(* IEC 61131-3 sources: SemaPLC/sema-plc-benchmark/spec2control-benchmark/data/st-baseline/paper-machine/pous/programs, 10 files *)

(* ---- main.st ---- *)
PROGRAM main
VAR
	Heartbeat : bool;
END_VAR

(* Entry point required by OpenPLC Editor v4. The process sections run as parallel program instances under task0; main only provides a scan heartbeat. *)
Heartbeat := NOT Heartbeat;

END_PROGRAM

(* ---- Section10.st ---- *)
PROGRAM Section10
VAR
	FT901_NipLoad_kN : real;
	FT902_FlowRate_Lmin : real;
	FIC904_Flow_SP_FromRatio : real;
	FT_901 : ANALOG_IN;
	FT_902 : ANALOG_IN;
	CW_901 : ANALOG_IN;
	FFIC_903 : RATIO_CONTROL;
	FIC_904 : PID_BASIC;
	FV_104 : VALVE_ELECTRIC;
	XV_105 : VALVE_ON_OFF;
	NipLoadOK_NOT : bool;
	SP_LowCut_SEL : real;
	XV105Closed_NOT : bool;
	CW901DevTrip_OR : bool;
	FT901_LowOrFault_OR : bool;
	CW901_DevOrFault_OR : bool;
	Interlock_PermissivesFail1_OR : bool;
	Interlock_PermissivesFail2_OR : bool;
	FFIC903_Inhibit_OR : bool;
END_VAR

FT_901(
    PV_Low := 5.0,
    Scaling_Slope := 6.25,
    Scaling_Offset := -25.0,
    Alarm_Enable := TRUE);
FT_902(
    Scaling_Slope := 31.25,
    Scaling_Offset := -125.0,
    Alarm_Enable := TRUE);
CW_901(
    Alarm_Enable := TRUE);
FT901_LowOrFault_OR := FT_901.Low_Alarm OR FT_901.General_Fault;
XV_105();
XV105Closed_NOT := NOT XV_105.FB_Opened;
Interlock_PermissivesFail1_OR := XV105Closed_NOT OR FT901_LowOrFault_OR;
CW901DevTrip_OR := CW_901.High_Alarm OR CW_901.Low_Alarm;
CW901_DevOrFault_OR := CW901DevTrip_OR OR CW_901.General_Fault;
Interlock_PermissivesFail2_OR := FT_902.General_Fault OR CW901_DevOrFault_OR;
FFIC903_Inhibit_OR := Interlock_PermissivesFail1_OR OR Interlock_PermissivesFail2_OR;
FFIC_903(
    Auto := TRUE,
    PrimaryPV := FT_901.PV,
    SecondaryPV := FT_902.PV,
    RatioSP := 2.0,
    Bias := 0.0,
    MV_MIN := 0.0,
    MV_MAX := 500.0,
    Inhibit := FFIC903_Inhibit_OR);
NipLoadOK_NOT := NOT FT_901.Low_Alarm;
SP_LowCut_SEL := SEL(G := NipLoadOK_NOT, IN0 := 0.0, IN1 := FFIC_903.SlaveSP);
FIC_904(
    AUTO := TRUE,
    PV := FT_902.PV,
    SP := SP_LowCut_SEL,
    MV_MIN := 0.0,
    MV_MAX := 100.0,
    X0 := 0.0,
    Deviation_Limit := 5.0);
FV_104(
    Control_Signal := FIC_904.XOUT,
    Manual_Mode := FALSE,
    Open_Limit := 100.0,
    Close_Limit := 0.0,
    Inhibit := FFIC903_Inhibit_OR);

(* Outputs published to other sections / HMI. *)
FT901_NipLoad_kN := FT_901.PV;
FT902_FlowRate_Lmin := FT_902.PV;
FIC904_Flow_SP_FromRatio := FFIC_903.SlaveSP;

END_PROGRAM

(* ---- Section2.st ---- *)
PROGRAM Section2
VAR
	LT_101_Flow_PV : real;
	FC_101_MV_to_FV106 : real;
	M_102_VSD_Speed_Out : real;
	Flow_Deviation_Alarm_30s : bool;
	Flow_High_Alarm : bool;
	Flow_Low_Alarm : bool;
	M_102_Start_Request : bool;
	M_102_Stop_Request : bool;
	LT_101 : ANALOG_IN;
	FC_101 : PID_BASIC;
	M_102 : MOTOR_VSD;
	FV_106 : VALVE_ELECTRIC;
	LV_103 : VALVE_ELECTRIC;
	XV_102 : VALVE_ON_OFF;
	XV_104 : VALVE_ON_OFF;
	XV_105 : VALVE_ON_OFF;
	FlowDeviationAlarm_TON : TON;
	M102_RestartDelay_TON : TON;
	FC101_ValvesOpen_AND : bool;
	FC101_ValvesNotOpen_NOT : bool;
	FC101_Inhibit_OR : bool;
	M102_XV105NotClosed_NOT : bool;
	M102_Inhibit_OR : bool;
	M102_InhibitNot_NOT : bool;
	M102_StartPermissive_AND : bool;
	M102_StopCmd_OR : bool;
	HopperLevelAbove20_GT : bool;
END_VAR

LT_101(
    PV_High := 380.0,
    PV_Low := 20.0,
    Scaling_Slope := 25.0,
    Scaling_Offset := -100.0,
    Alarm_Enable := TRUE);
XV_105(
    Timeout := T#5s);
M102_XV105NotClosed_NOT := NOT XV_105.FB_Closed;
M102_Inhibit_OR := M102_XV105NotClosed_NOT OR LT_101.General_Fault;
LV_103(
    Open_Limit := 100.0,
    Close_Limit := 0.0);
HopperLevelAbove20_GT := (LV_103.Feedback_Pos > 20.0);
M102_InhibitNot_NOT := NOT M102_Inhibit_OR;
M102_RestartDelay_TON(
    IN := M102_InhibitNot_NOT,
    PT := T#60s);
M102_StartPermissive_AND := HopperLevelAbove20_GT AND XV_105.FB_Closed AND M102_RestartDelay_TON.Q AND M_102_Start_Request;
M102_StopCmd_OR := M_102_Stop_Request OR M102_Inhibit_OR;
M_102(
    Start_Cmd := M102_StartPermissive_AND,
    Stop_Cmd := M102_StopCmd_OR,
    Accel_Ramp := T#2s,
    Decel_Ramp := T#2s,
    Inhibit := M102_Inhibit_OR);
XV_102(
    Timeout := T#5s,
    Inhibit := M_102.FB_Fault);
XV_104(
    Timeout := T#5s,
    Inhibit := M_102.FB_Fault);
FC101_ValvesOpen_AND := XV_102.FB_Opened AND XV_104.FB_Opened;
FC101_ValvesNotOpen_NOT := NOT FC101_ValvesOpen_AND;
FC101_Inhibit_OR := FC101_ValvesNotOpen_NOT OR LT_101.General_Fault OR M_102.FB_Fault;
FC_101(
    AUTO := TRUE,
    PV := LT_101.PV,
    SP := 250.0,
    MV_MIN := 0.0,
    MV_MAX := 100.0,
    KP := 3.0,
    TR := 1.2,
    TD := 0.3,
    Deviation_Limit := 5.0,
    Inhibit := FC101_Inhibit_OR);
FV_106(
    Control_Signal := FC_101.XOUT,
    Manual_Mode := FALSE,
    Manual_Position := 0.0,
    Open_Limit := 100.0,
    Close_Limit := 0.0,
    Timeout := T#5s,
    Inhibit := LT_101.General_Fault);
FlowDeviationAlarm_TON(
    IN := FC_101.Deviation_Alarm,
    PT := T#30s);

(* Outputs published to other sections / HMI. *)
FC_101_MV_to_FV106 := FC_101.XOUT;
LT_101_Flow_PV := LT_101.PV;
Flow_High_Alarm := LT_101.High_Alarm;
Flow_Low_Alarm := LT_101.Low_Alarm;
Flow_Deviation_Alarm_30s := FlowDeviationAlarm_TON.Q;
M_102_VSD_Speed_Out := M_102.Speed_Out;

END_PROGRAM

(* ---- Section3.st ---- *)
PROGRAM Section3
VAR
	TT_103_Temperature_PV : real;
	PT_101_Pressure_PV : real;
	TIC_104_RSP_to_FC_203 : real;
	PIC_101_RSP_to_FC_202 : real;
	FC_203_MV_to_SV_203 : real;
	FC_202_MV_to_FV_202 : real;
	TT_103 : ANALOG_IN;
	PT_101 : ANALOG_IN;
	TIC_104 : PID_BASIC;
	PIC_101 : PID_BASIC;
	FC_203 : PID_BASIC;
	FC_202 : PID_BASIC;
	SV_203 : VALVE_ELECTRIC;
	FV_202 : VALVE_ELECTRIC;
	SV203Trip_OR : bool;
	CascadeInhibit_OR : bool;
END_VAR

TT_103(
    PV_High := 180.0,
    PV_Low := 160.0,
    Scaling_Slope := 11.25,
    Scaling_Offset := -25.0,
    Alarm_Enable := TRUE);
PT_101(
    Alarm_Enable := TRUE);
PIC_101(
    AUTO := TRUE,
    PV := PT_101.PV,
    SP := 800.0,
    MV_MIN := 0.0,
    MV_MAX := 100.0,
    PV_High := 850.0,
    PV_Low := 750.0,
    Inhibit := CascadeInhibit_OR);
FC_202(
    AUTO := TRUE,
    SP := PIC_101.XOUT,
    MV_MIN := 0.0,
    MV_MAX := 100.0,
    Inhibit := PIC_101.PV_Low_Alarm);
FV_202(
    Control_Signal := FC_202.XOUT);
FC_203(
    AUTO := TRUE,
    SP := TIC_104.XOUT,
    MV_MIN := 0.0,
    MV_MAX := 100.0,
    KP := 3.5,
    TR := 0.3,
    Inhibit := TT_103.General_Fault);
SV203Trip_OR := PIC_101.PV_High_Alarm OR TIC_104.PV_High_Alarm;
SV_203(
    Control_Signal := FC_203.XOUT,
    Inhibit := SV203Trip_OR);
CascadeInhibit_OR := TT_103.General_Fault OR PT_101.General_Fault OR SV_203.Alarm OR FV_202.Alarm;
TIC_104(
    AUTO := TRUE,
    PV := TT_103.PV,
    SP := 170.0,
    MV_MIN := 0.0,
    MV_MAX := 100.0,
    KP := 1.2,
    TR := 2.0,
    Inhibit := CascadeInhibit_OR);

(* Outputs published to other sections / HMI. *)
TT_103_Temperature_PV := TT_103.PV;
PT_101_Pressure_PV := PT_101.PV;
TIC_104_RSP_to_FC_203 := TIC_104.XOUT;
PIC_101_RSP_to_FC_202 := PIC_101.XOUT;
FC_203_MV_to_SV_203 := FC_203.XOUT;
FC_202_MV_to_FV_202 := FC_202.XOUT;

END_PROGRAM

(* ---- Section4.st ---- *)
PROGRAM Section4
VAR
	PIT103_Pressure_kPa : real;
	PT101_UpstreamPressure_kPa : real;
	DT301_PulpDensity_Pct : real;
	PIC104_ControlOutput_to_FV106_Pct : real;
	FV106_ValvePositionFeedback_Pct : real;
	DT_301 : ANALOG_IN;
	PIT_103 : ANALOG_IN;
	PT_101 : ANALOG_IN;
	PIC_104 : PID_BASIC;
	FV_106 : VALVE_ELECTRIC;
	XV_102 : VALVE_ON_OFF;
	XV_107 : VALVE_ON_OFF;
	XV_102_OPEN_FB : DIGITAL_IN;
	XV_107_OPEN_FB : DIGITAL_IN;
	PERM_XV102_OPEN : BOOL_INPUT;
	PERM_XV107_OPEN : BOOL_INPUT;
	PIC104Inhibit_OR : bool;
	FV106Inhibit_OR : bool;
	SystemFault_OR : bool;
	XV102NotOpen_NOT : bool;
	XV107NotOpen_NOT : bool;
	SystemEnable_NOT : bool;
	PIC104Auto_NOT : bool;
END_VAR

DT_301();
PIT_103(
    Scaling_Slope := 31.25,
    Scaling_Offset := -125.0);
PT_101();
PIC104Inhibit_OR := PT_101.Low_Alarm OR PT_101.High_Alarm OR DT_301.High_Alarm OR PIT_103.General_Fault;
PIC104Auto_NOT := NOT PIC104Inhibit_OR;
PIC_104(
    AUTO := PIC104Auto_NOT,
    PV := PIT_103.PV,
    SP := 250.0,
    MV_MIN := 0.0,
    MV_MAX := 100.0,
    X0 := 0.0,
    KP := -3.0,
    TR := 1.2,
    TD := 0.1,
    PV_High := 275.0,
    PV_Low := 200.0,
    Deviation_Limit := 12.5,
    Inhibit := PIC104Inhibit_OR);
XV_102_OPEN_FB();
PERM_XV102_OPEN(
    Bool_In := XV_102_OPEN_FB.DI_Out);
XV102NotOpen_NOT := NOT PERM_XV102_OPEN.Bool_Out;
XV_107_OPEN_FB();
PERM_XV107_OPEN(
    Bool_In := XV_107_OPEN_FB.DI_Out);
XV107NotOpen_NOT := NOT PERM_XV107_OPEN.Bool_Out;
FV106Inhibit_OR := XV102NotOpen_NOT OR XV107NotOpen_NOT OR PT_101.High_Alarm OR PIT_103.General_Fault;
FV_106(
    Control_Signal := PIC_104.XOUT,
    Manual_Mode := FALSE,
    Manual_Position := 0.0,
    Open_Limit := 100.0,
    Close_Limit := 0.0,
    Timeout := T#2S,
    Inhibit := FV106Inhibit_OR);
SystemFault_OR := PT_101.General_Fault OR DT_301.General_Fault;
SystemEnable_NOT := NOT SystemFault_OR;
XV_102(
    Open_Cmd := SystemEnable_NOT,
    Close_Cmd := SystemFault_OR,
    Inhibit := SystemFault_OR);
XV_107(
    Open_Cmd := SystemEnable_NOT,
    Close_Cmd := SystemFault_OR,
    Inhibit := SystemFault_OR);

(* Outputs published to other sections / HMI. *)
PIT103_Pressure_kPa := PIT_103.PV;
PT101_UpstreamPressure_kPa := PT_101.PV;
DT301_PulpDensity_Pct := DT_301.PV;
PIC104_ControlOutput_to_FV106_Pct := PIC_104.XOUT;
FV106_ValvePositionFeedback_Pct := FV_106.Feedback_Pos;

END_PROGRAM

(* ---- Section5.st ---- *)
PROGRAM Section5
VAR
	AT102_pH_PV : real;
	AT107_pH_PV : real;
	TIT106_Temperature_PV : real;
	LIC102_MV_to_FV101 : real;
	TIC106_MV_to_FV103 : real;
	LIC104_MV_to_XV104 : real;
	AT_102 : ANALOG_IN;
	AT_107 : ANALOG_IN;
	TIT_106 : ANALOG_IN;
	LIC_102 : PID_BASIC;
	TIC_106 : PID_BASIC;
	LIC_104 : PID_BASIC;
	FV_101 : VALVE_ELECTRIC;
	FV_103 : VALVE_ELECTRIC;
	XV_104 : VALVE_ELECTRIC;
	PHExtremeTrip_OR : bool;
END_VAR

AT_102(
    Scaling_Slope := 0.875,
    Scaling_Offset := -3.5,
    Alarm_Enable := TRUE);
AT_107(
    Alarm_Enable := TRUE);
TIT_106(
    Scaling_Slope := 6.25,
    Scaling_Offset := -25.0,
    Alarm_Enable := TRUE);
FV_101(
    Control_Signal := LIC_102.XOUT,
    Open_Limit := 100.0,
    Close_Limit := 0.0,
    Timeout := T#10s,
    Inhibit := AT_107.General_Fault);
PHExtremeTrip_OR := LIC_102.PV_High_Alarm OR LIC_102.PV_Low_Alarm;
LIC_102(
    AUTO := TRUE,
    PV := AT_102.PV,
    SP := 9.25,
    MV_MIN := 10.0,
    MV_MAX := 90.0,
    X0 := FV_101.Feedback_Pos,
    KP := 1.8,
    TR := 0.5,
    TD := 0.1,
    PV_High := 10.5,
    PV_Low := 8.5,
    Deviation_Limit := 1.0,
    Inhibit := PHExtremeTrip_OR);
FV_103(
    Control_Signal := TIC_106.XOUT,
    Open_Limit := 100.0,
    Close_Limit := 0.0,
    Timeout := T#10s);
TIC_106(
    AUTO := TRUE,
    PV := TIT_106.PV,
    SP := 65.0,
    MV_MIN := 0.0,
    MV_MAX := 100.0,
    X0 := FV_103.Feedback_Pos,
    KP := 2.0,
    TR := 0.4,
    TD := 0.05,
    PV_High := 75.0,
    PV_Low := 55.0,
    Inhibit := TIC_106.PV_High_Alarm);
XV_104(
    Control_Signal := LIC_104.XOUT,
    Open_Limit := 100.0,
    Close_Limit := 0.0,
    Timeout := T#10s);
LIC_104(
    AUTO := TRUE,
    SP := 120.0,
    MV_MIN := 0.0,
    MV_MAX := 100.0,
    X0 := XV_104.Feedback_Pos,
    KP := 1.5,
    TR := 1.0,
    TD := 0.2,
    Deviation_Limit := 10.0);

(* Outputs published to other sections / HMI. *)
AT102_pH_PV := AT_102.PV;
AT107_pH_PV := AT_107.PV;
TIT106_Temperature_PV := TIT_106.PV;
LIC102_MV_to_FV101 := LIC_102.XOUT;
TIC106_MV_to_FV103 := TIC_106.XOUT;
LIC104_MV_to_XV104 := LIC_104.XOUT;

END_PROGRAM

(* ---- Section6.st ---- *)
PROGRAM Section6
VAR
	CT501_Consistency_PV_Pct : real;
	FC502_MV_to_FV502_Pct : real;
	SELT501_SEL_PV_WsPerMm2 : real;
	SELC501_MV_to_PGA501_Pct : real;
	LT501_Level_PV_Pct : real;
	PT502_Pressure_PV_kPa : real;
	PGT501_PlateGap_PV_mm : real;
	CT_501 : ANALOG_IN;
	FC_502 : PID_BASIC;
	FV_502 : VALVE_ELECTRIC;
	LT_501 : ANALOG_IN;
	M_501 : MOTOR_ON_OFF;
	PT_502 : ANALOG_IN;
	SELC_501 : PID_BASIC;
	PGT_501 : ANALOG_IN;
	PGA_501 : VALVE_ELECTRIC;
	SELT_501 : ANALOG_IN;
	INTLK_M501_RUNNING : BOOL_INPUT;
	INTLK_PLATE_GAP_IN_RANGE : BOOL_INPUT;
	INTLK_LEVEL_ABOVE_20 : BOOL_INPUT;
	PERM_PT502_IN_RANGE : BOOL_INPUT;
	PGT501_OutOfRange_OR : bool;
	PlateGapInRange_NOT : bool;
	SEL_Enable_AND : bool;
	SEL_Inhibit_NOT : bool;
	LT501_LevelNotOK_OR : bool;
	LevelAbove20_NOT : bool;
	PT502_NotInRange_OR : bool;
	PT502_InRange_NOT : bool;
	FC502_Inhibit_OR : bool;
END_VAR

CT_501(
    Scaling_Slope := 0.1875,
    Scaling_Offset := 1.25,
    Alarm_Enable := TRUE);
LT_501(
    Alarm_Enable := TRUE);
LT501_LevelNotOK_OR := LT_501.Low_Alarm OR LT_501.General_Fault;
PT_502(
    Alarm_Enable := TRUE);
PT502_NotInRange_OR := PT_502.High_Alarm OR PT_502.Low_Alarm OR PT_502.General_Fault;
FC502_Inhibit_OR := LT501_LevelNotOK_OR OR PT502_NotInRange_OR OR CT_501.General_Fault;
FC_502(
    AUTO := TRUE,
    PV := CT_501.PV,
    SP := 3.0,
    MV_MIN := 0.0,
    MV_MAX := 100.0,
    X0 := 0.0,
    KP := 2.2,
    TR := 0.7,
    TD := 0.0,
    PV_High := 4.0,
    PV_Low := 2.0,
    Inhibit := FC502_Inhibit_OR);
FV_502(
    Control_Signal := FC_502.XOUT,
    Manual_Mode := FALSE,
    Open_Limit := 100.0,
    Close_Limit := 0.0,
    Inhibit := FC502_Inhibit_OR);
PGT_501(
    Alarm_Enable := TRUE);
PGT501_OutOfRange_OR := PGT_501.High_Alarm OR PGT_501.Low_Alarm OR PGT_501.General_Fault;
M_501(
    Inhibit := PGT501_OutOfRange_OR);
SELT_501(
    Scaling_Slope := 0.0625,
    Scaling_Offset := -0.05,
    Alarm_Enable := TRUE);
INTLK_M501_RUNNING(
    Bool_In := M_501.FB_Running);
PlateGapInRange_NOT := NOT PGT501_OutOfRange_OR;
INTLK_PLATE_GAP_IN_RANGE(
    Bool_In := PlateGapInRange_NOT);
SEL_Enable_AND := INTLK_M501_RUNNING.Bool_Out AND INTLK_PLATE_GAP_IN_RANGE.Bool_Out;
SEL_Inhibit_NOT := NOT SEL_Enable_AND;
SELC_501(
    AUTO := TRUE,
    PV := SELT_501.PV,
    MV_MIN := 0.0,
    MV_MAX := 100.0,
    X0 := 0.0,
    KP := 1.8,
    TR := 0.5,
    TD := 0.1,
    PV_High := 1.1,
    PV_Low := 0.3,
    Inhibit := SEL_Inhibit_NOT);
PGA_501(
    Control_Signal := SELC_501.XOUT,
    Manual_Mode := FALSE,
    Open_Limit := 100.0,
    Close_Limit := 0.0);
LevelAbove20_NOT := NOT LT501_LevelNotOK_OR;
INTLK_LEVEL_ABOVE_20(
    Bool_In := LevelAbove20_NOT);
PT502_InRange_NOT := NOT PT502_NotInRange_OR;
PERM_PT502_IN_RANGE(
    Bool_In := PT502_InRange_NOT);

(* Outputs published to other sections / HMI. *)
CT501_Consistency_PV_Pct := CT_501.PV;
FC502_MV_to_FV502_Pct := FC_502.XOUT;
SELT501_SEL_PV_WsPerMm2 := SELT_501.PV;
SELC501_MV_to_PGA501_Pct := SELC_501.XOUT;
LT501_Level_PV_Pct := LT_501.PV;
PT502_Pressure_PV_kPa := PT_502.PV;
PGT501_PlateGap_PV_mm := PGT_501.PV;

END_PROGRAM

(* ---- Section7.st ---- *)
PROGRAM Section7
VAR
	CT_601_PV : real;
	FT_601_PV : real;
	FT_601_SP : real;
	PIT_601_PV : real;
	VT_601_PV : real;
	FS_601_MinFlow_OK : bool;
	P_601_Run_OK : bool;
	FFIC601_Bias : real;
	ALM_601 : bool;
	ALM_601_High : bool;
	ALM_601_Low : bool;
	ALM_602 : bool;
	ALM_603 : bool;
	ALM_604 : bool;
	Process_Permissives_OK : bool;
	MasterInhibit : bool;
	CT601_RateHigh : bool;
	CT_601 : ANALOG_IN;
	FT_601 : ANALOG_IN;
	PIT_601 : ANALOG_IN;
	VT_601 : ANALOG_IN;
	FS_601 : BOOL_INPUT;
	P_601_RUN : BOOL_INPUT;
	FV_601 : VALVE_ELECTRIC;
	FIC_601 : PID_BASIC;
	FFIC_601 : RATIO_CONTROL;
	ProcessUpset_Timer : TON;
	PumpRun_Fault : bool;
	MinFlow_Fault : bool;
	CT_Failure : bool;
	FT_Failure : bool;
	Inhibit_Any : bool;
	Auto_Enable : bool;
	SlaveSP_TooHigh : bool;
	SlaveSP_TooLow : bool;
	SlaveSP_LimitAlarm : bool;
END_VAR

CT_601(
    Alarm_Enable := TRUE);
FT_601(
    PV_High := 500.0,
    PV_Low := 10.0,
    Alarm_Enable := TRUE);
PIT_601(
    PV_Low := 300.0,
    Alarm_Enable := TRUE);
VT_601(
    Alarm_Enable := TRUE);
FS_601(
    Alarm_OnFalse := TRUE);
P_601_RUN(
    Alarm_OnFalse := TRUE);
CT_Failure := CT_601.High_Alarm OR CT_601.Low_Alarm OR CT_601.General_Fault;
FT_Failure := FT_601.High_Alarm OR FT_601.Low_Alarm OR FT_601.General_Fault;
MinFlow_Fault := NOT FS_601.Bool_Out;
PumpRun_Fault := NOT P_601_RUN.Bool_Out;
Inhibit_Any := PumpRun_Fault OR MinFlow_Fault OR PIT_601.Low_Alarm OR VT_601.Low_Alarm OR CT_Failure OR FT_Failure;
Auto_Enable := NOT Inhibit_Any;
FFIC_601(
    Auto := Auto_Enable,
    PrimaryPV := CT_601.PV,
    SecondaryPV := FT_601.PV,
    RatioSP := 2.5,
    Bias := FFIC601_Bias,
    TrimKp := 0.1,
    TrimTi := T#2s,
    MV_MIN := 10.0,
    MV_MAX := 500.0,
    Inhibit := Inhibit_Any);
FIC_601(
    AUTO := Auto_Enable,
    PV := FT_601.PV,
    SP := FFIC_601.SlaveSP,
    MV_MIN := 0.0,
    MV_MAX := 100.0,
    X0 := 20.0,
    Inhibit := Inhibit_Any);
FV_601(
    Control_Signal := FIC_601.XOUT,
    Manual_Mode := Inhibit_Any,
    Manual_Position := 20.0,
    Open_Limit := 100.0,
    Close_Limit := 0.0,
    Inhibit := Inhibit_Any);
ProcessUpset_Timer(
    IN := CT601_RateHigh,
    PT := T#10s);
SlaveSP_TooHigh := (FFIC_601.SlaveSP > 500.0);
SlaveSP_TooLow := (FFIC_601.SlaveSP < 10.0);
SlaveSP_LimitAlarm := SlaveSP_TooHigh OR SlaveSP_TooLow;

(* Outputs published to other sections / HMI. *)
ALM_601 := SlaveSP_LimitAlarm;
ALM_602 := CT_Failure;
ALM_603 := FT_Failure;
ALM_604 := ProcessUpset_Timer.Q;
CT_601_PV := CT_601.PV;
FT_601_PV := FT_601.PV;
FT_601_SP := FFIC_601.SlaveSP;
PIT_601_PV := PIT_601.PV;
VT_601_PV := VT_601.PV;
FS_601_MinFlow_OK := FS_601.Bool_Out;
P_601_Run_OK := P_601_RUN.Bool_Out;
MasterInhibit := Inhibit_Any;
Process_Permissives_OK := Auto_Enable;

END_PROGRAM

(* ---- Section8.st ---- *)
PROGRAM Section8
VAR
	MM701_Raw_mA : real;
	PT701_Raw : real;
	TT102_Raw : real;
	HS701_ON : bool;
	CS701_ON : bool;
	SB701_SheetBreak : bool;
	MM701_Moisture_PV : real;
	PT701_HydraulicPressure_PV : real;
	TT102_ShowerWaterTemp_PV : real;
	PV101_Pressure_Command_Pct : real;
	PV101_Position_Feedback_Pct : real;
	ESD_Trip : bool;
	MM_701 : ANALOG_IN;
	PT_701 : ANALOG_IN;
	TT_102 : ANALOG_IN;
	LIC_701 : PID_BASIC;
	PV_101 : VALVE_ELECTRIC;
	HS_701 : BOOL_INPUT;
	CS_701 : BOOL_INPUT;
	SB_701 : BOOL_INPUT;
	SheetPresent_NOT : bool;
	PressLoopPermissive_AND : bool;
	FailCloseTrip_OR : bool;
	LoopInhibit_OR : bool;
	MoistureTrip_GT : bool;
END_VAR

MM_701(
    Raw_Signal := MM701_Raw_mA,
    PV_High := 58.0,
    PV_Low := 46.0,
    Scaling_Slope := 1.25,
    Scaling_Offset := 35.0,
    Alarm_Enable := TRUE);
PT_701(
    Raw_Signal := PT701_Raw,
    Scaling_Slope := 1.0,
    Scaling_Offset := 0.0,
    Alarm_Enable := TRUE);
TT_102(
    Raw_Signal := TT102_Raw,
    Scaling_Slope := 1.0,
    Scaling_Offset := 0.0,
    Alarm_Enable := TRUE);
MoistureTrip_GT := (MM_701.PV > 65.0);
PV_101(
    Control_Signal := LIC_701.XOUT,
    Manual_Mode := FailCloseTrip_OR,
    Manual_Position := 0.0,
    Open_Limit := 100.0,
    Close_Limit := 0.0);
FailCloseTrip_OR := TT_102.High_Alarm OR MoistureTrip_GT OR PT_701.High_Alarm OR PV_101.Position_Error;
LoopInhibit_OR := MM_701.General_Fault OR FailCloseTrip_OR;
CS_701(
    Bool_In := CS701_ON);
HS_701(
    Bool_In := HS701_ON);
SB_701(
    Bool_In := SB701_SheetBreak);
SheetPresent_NOT := NOT SB_701.Bool_Out;
PressLoopPermissive_AND := HS_701.Bool_Out AND CS_701.Bool_Out AND SheetPresent_NOT;
LIC_701(
    AUTO := PressLoopPermissive_AND,
    PV := MM_701.PV,
    SP := 52.0,
    MV_MIN := 0.0,
    MV_MAX := 100.0,
    X0 := PV_101.Feedback_Pos,
    KP := 3.0,
    TR := 1.2,
    TD := 0.2,
    Deviation_Limit := 2.0,
    Inhibit := LoopInhibit_OR);

(* Outputs published to other sections / HMI. *)
MM701_Moisture_PV := MM_701.PV;
PT701_HydraulicPressure_PV := PT_701.PV;
TT102_ShowerWaterTemp_PV := TT_102.PV;
PV101_Pressure_Command_Pct := LIC_701.XOUT;
PV101_Position_Feedback_Pct := PV_101.Feedback_Pos;
ESD_Trip := PT_701.High_Alarm;

END_PROGRAM

(* ---- Section9.st ---- *)
PROGRAM Section9
VAR
	F801_ExhaustFan_Speed_CMD_PCT : real;
	FV801_SteamFlowValve_Position_CMD_PCT : real;
	XV802_HotAirDamper_Position_CMD_PCT : real;
	WT801_DownstreamDriveRoll_Torque_CMD_PCT : real;
	XV802_Open_FB : bool;
	IR801_Available : bool;
	TT_801 : ANALOG_IN;
	TT_802 : ANALOG_IN;
	PT_801 : ANALOG_IN;
	IR_801 : ANALOG_IN;
	WT_801 : ANALOG_IN;
	F_801 : MOTOR_VSD;
	M_801 : MOTOR_ON_OFF;
	FV_801 : VALVE_ELECTRIC;
	XV_802 : VALVE_ELECTRIC;
	SC_801 : PID_BASIC;
	TC_801 : PID_BASIC;
	F_801_CTRL : PID_BASIC;
	WT_801_CTRL : PID_BASIC;
	SteamFlowInterlock : bool;
	XV802NotOpen : bool;
	HoodTempInhibit : bool;
	IR801NotAvailable : bool;
	FanControlInhibit : bool;
	M801NotRunning : bool;
	WebTensionInhibit : bool;
	DriveStop : bool;
END_VAR

TT_801(
    Scaling_Slope := 9.375,
    Scaling_Offset := -37.5,
    Alarm_Enable := TRUE);
TT_802(
    Scaling_Slope := 4.375,
    Scaling_Offset := 32.5,
    Alarm_Enable := TRUE);
PT_801(
    PV_Low := 600.0,
    Alarm_Enable := TRUE);
IR_801(
    PV_High := 5.0,
    Scaling_Slope := 0.625,
    Scaling_Offset := -2.5,
    Alarm_Enable := TRUE);
WT_801(
    Scaling_Slope := 31.25,
    Scaling_Offset := -125.0,
    Alarm_Enable := TRUE);
IR801NotAvailable := NOT IR801_Available;
FanControlInhibit := IR801NotAvailable OR IR_801.High_Alarm OR IR_801.Low_Alarm OR IR_801.General_Fault;
F_801_CTRL(
    AUTO := TRUE,
    PV := IR_801.PV,
    SP := 4.5,
    MV_MIN := 0.0,
    MV_MAX := 100.0,
    KP := 1.8,
    TR := 0.6,
    TD := 0.05,
    Deviation_Limit := 0.2,
    Inhibit := FanControlInhibit);
F_801(
    Speed_SP := F_801_CTRL.XOUT,
    Inhibit := FanControlInhibit);
DriveStop := WT_801.High_Alarm OR WT_801.Low_Alarm;
M_801(
    Inhibit := DriveStop);
SteamFlowInterlock := PT_801.High_Alarm OR PT_801.Low_Alarm OR SC_801.PV_High_Alarm;
SC_801(
    AUTO := TRUE,
    PV := TT_801.PV,
    SP := 115.0,
    MV_MIN := 0.0,
    MV_MAX := 100.0,
    KP := 3.0,
    TR := 0.5,
    TD := 0.1,
    PV_High := 125.0,
    Inhibit := SteamFlowInterlock);
FV_801(
    Control_Signal := SC_801.XOUT,
    Open_Limit := 100.0,
    Close_Limit := 0.0,
    Inhibit := SteamFlowInterlock);
XV802NotOpen := NOT XV802_Open_FB;
HoodTempInhibit := XV802NotOpen OR TT_802.High_Alarm OR TT_802.Low_Alarm;
TC_801(
    AUTO := TRUE,
    PV := TT_802.PV,
    SP := 85.0,
    MV_MIN := 10.0,
    MV_MAX := 90.0,
    KP := 2.5,
    TR := 0.8,
    TD := 0.2,
    PV_High := 95.0,
    Inhibit := HoodTempInhibit);
XV_802(
    Control_Signal := TC_801.XOUT,
    Open_Limit := 90.0,
    Close_Limit := 10.0,
    Inhibit := TC_801.PV_High_Alarm);
M801NotRunning := NOT M_801.FB_Running;
WebTensionInhibit := M801NotRunning OR WT_801.High_Alarm OR WT_801.Low_Alarm;
WT_801_CTRL(
    AUTO := TRUE,
    PV := WT_801.PV,
    SP := 250.0,
    MV_MIN := 0.0,
    MV_MAX := 100.0,
    KP := 4.0,
    TR := 1.0,
    TD := 0.3,
    PV_High := 400.0,
    Inhibit := WebTensionInhibit);

(* Outputs published to other sections / HMI. *)
WT801_DownstreamDriveRoll_Torque_CMD_PCT := WT_801_CTRL.XOUT;
F801_ExhaustFan_Speed_CMD_PCT := F_801.Speed_Out;
FV801_SteamFlowValve_Position_CMD_PCT := FV_801.Valve_Position;
XV802_HotAirDamper_Position_CMD_PCT := XV_802.Valve_Position;

END_PROGRAM
